(* IEC 61131-3 sources: trust-platform/examples/OSCAT/temperature_zone_composition/non-oop/src, 3 files *)

(* ---- Configuration.st ---- *)
CONFIGURATION TemperatureZoneCompositionClassicConfiguration
RESOURCE TemperatureZoneCompositionClassic ON PLC
    TASK MainTask (INTERVAL := T#100ms, PRIORITY := 1);
    PROGRAM Main WITH MainTask : Main;
END_RESOURCE
END_CONFIGURATION

(* ---- Main.st ---- *)
PROGRAM Main
VAR
    ZoneAFilter : FT_PT1;
    ZoneBFilter : FT_PT1;
    ZoneAController : CTRL_PID;
    ZoneBController : CTRL_PID;
    ZoneAAlarm : HYST;
    ZoneBAlarm : HYST;
    ZoneACommand : REAL;
    ZoneBCommand : REAL;
    AnyAlarm : BOOL;
END_VAR

ZoneAFilter(in := REAL#21.0, T := T#1s, K := REAL#1.0);
ZoneAController(ACT := ZoneAFilter.out, SET_POINT := REAL#23.0, SUP := REAL#0.0, OFS := REAL#0.0, M_I := REAL#45.0, MAN := TRUE, RST := FALSE, KP := REAL#1.0, TN := REAL#1.0, TV := REAL#0.0, LL := REAL#0.0, LH := REAL#100.0);
ZoneAAlarm(In := ZoneAFilter.out, HIGH_LIMIT := REAL#30.0, LOW_LIMIT := REAL#5.0);
ZoneACommand := ZoneAController.Y;

ZoneBFilter(in := REAL#18.0, T := T#1s, K := REAL#1.0);
ZoneBController(ACT := ZoneBFilter.out, SET_POINT := REAL#22.0, SUP := REAL#0.0, OFS := REAL#0.0, M_I := REAL#55.0, MAN := TRUE, RST := FALSE, KP := REAL#1.0, TN := REAL#1.0, TV := REAL#0.0, LL := REAL#0.0, LH := REAL#100.0);
ZoneBAlarm(In := ZoneBFilter.out, HIGH_LIMIT := REAL#30.0, LOW_LIMIT := REAL#5.0);
ZoneBCommand := ZoneBController.Y;

AnyAlarm := ZoneAAlarm.Q OR ZoneBAlarm.Q;
END_PROGRAM

(* ---- Tests.st ---- *)
TEST_PROGRAM TemperatureZoneClassicRepeatsTheThreeBlockPattern
VAR
    ZoneFilter : FT_PT1;
    ZoneController : CTRL_PID;
    ZoneAlarm : HYST;
END_VAR

ZoneFilter(in := REAL#21.0, T := T#1s, K := REAL#1.0);
ZoneController(ACT := ZoneFilter.out, SET_POINT := REAL#23.0, SUP := REAL#0.0, OFS := REAL#0.0, M_I := REAL#45.0, MAN := TRUE, RST := FALSE, KP := REAL#1.0, TN := REAL#1.0, TV := REAL#0.0, LL := REAL#0.0, LH := REAL#100.0);
ZoneAlarm(In := ZoneFilter.out, HIGH_LIMIT := REAL#30.0, LOW_LIMIT := REAL#5.0);

ASSERT_NEAR(EXPECTED := REAL#21.0, ACTUAL := ZoneFilter.out, DELTA := REAL#0.001);
ASSERT_NEAR(EXPECTED := REAL#45.0, ACTUAL := ZoneController.Y, DELTA := REAL#0.001);
ASSERT_FALSE(IN := ZoneAlarm.Q);
END_TEST_PROGRAM
